(* IEC 61131-3 sources: llm-plc-st-eval/data/definitivo/gpt-4o-2024-08-06/I8/few_shot, 3 files *)

(* ---- ejec_1.st ---- *)
```pascal
FUNCTION_BLOCK FB_Compresor
VAR_INPUT
    pOilOk : BOOL; (* Presión de aceite correcta *)
    tempOk : BOOL; (* Temperatura correcta *)
    sinAlm : BOOL; (* Ausencia de alarmas *)
    btnMarcha : BOOL; (* Botón de marcha *)
    btnParo : BOOL; (* Botón de paro *)
END_VAR
VAR_OUTPUT
    comp : BOOL; (* Compresor en marcha *)
    causaBloqueo : INT; (* Causa de bloqueo *)
END_VAR
VAR
    pOilOkTimer : TON; (* Temporizador para presión de aceite *)
    btnMarchaMem : BOOL; (* Memoria del estado del botón de marcha *)
    btnMarchaRising : BOOL; (* Detección de flanco ascendente del botón de marcha *)
END_VAR

(* Detección de flanco ascendente del botón de marcha *)
btnMarchaRising := btnMarcha AND NOT btnMarchaMem;
btnMarchaMem := btnMarcha;

(* Temporizador para verificar presión de aceite durante 3 segundos continuos *)
pOilOkTimer(IN := pOilOk, PT := T#3S);

(* Determinación de la causa de bloqueo *)
IF NOT pOilOkTimer.Q THEN
    causaBloqueo := 1; (* Falta presión de aceite *)
ELSIF NOT tempOk THEN
    causaBloqueo := 2; (* Falta temperatura correcta *)
ELSIF NOT sinAlm THEN
    causaBloqueo := 3; (* Alarma activa *)
ELSE
    causaBloqueo := 0; (* Ningún bloqueo *)
END_IF

(* Lógica de control del compresor *)
IF btnParo THEN
    comp := FALSE; (* Parar compresor si se pulsa el botón de paro *)
ELSIF comp THEN
    IF causaBloqueo <> 0 THEN
        comp := FALSE; (* Parar compresor si se pierde algún permisivo *)
    END_IF
ELSE
    IF btnMarchaRising AND (causaBloqueo = 0) THEN
        comp := TRUE; (* Arrancar compresor si se pulsa el botón de marcha y no hay bloqueos *)
    END_IF
END_IF

END_FUNCTION_BLOCK
```

(* ---- ejec_2.st ---- *)
```pascal
FUNCTION_BLOCK FB_Compresor
VAR_INPUT
    pOilOk : BOOL; (* Presion de aceite correcta *)
    tempOk : BOOL; (* Temperatura correcta *)
    sinAlm : BOOL; (* Ausencia de alarmas *)
    btnMarcha : BOOL; (* Boton de marcha *)
    btnParo : BOOL; (* Boton de paro *)
END_VAR
VAR_OUTPUT
    comp : BOOL; (* Compresor en marcha *)
    causaBloqueo : INT; (* Causa de bloqueo *)
END_VAR
VAR
    pOilOkTimer : TON; (* Temporizador para presion de aceite *)
    btnMarchaMem : BOOL; (* Memoria de estado del boton de marcha *)
    permisivosOk : BOOL; (* Todos los permisivos estan activos *)
END_VAR

(* Temporizador para verificar presion de aceite durante 3 segundos *)
pOilOkTimer(IN := pOilOk, PT := T#3S);

(* Verificar si todos los permisivos estan activos *)
permisivosOk := pOilOkTimer.Q AND tempOk AND sinAlm;

(* Logica de arranque y paro del compresor *)
IF btnParo THEN
    comp := FALSE; (* Parar compresor si se pulsa btnParo *)
ELSIF NOT comp AND NOT btnMarchaMem AND btnMarcha AND permisivosOk THEN
    comp := TRUE; (* Arrancar compresor si se pulsa btnMarcha y permisivos estan activos *)
END_IF

(* Actualizar memoria del estado del boton de marcha *)
btnMarchaMem := btnMarcha;

(* Determinar la causa de bloqueo *)
IF NOT pOilOk THEN
    causaBloqueo := 1; (* Bloqueo por presion de aceite *)
ELSIF NOT tempOk THEN
    causaBloqueo := 2; (* Bloqueo por temperatura *)
ELSIF NOT sinAlm THEN
    causaBloqueo := 3; (* Bloqueo por alarma activa *)
ELSE
    causaBloqueo := 0; (* No hay bloqueo *)
END_IF
END_FUNCTION_BLOCK
```

(* ---- ejec_3.st ---- *)
```pascal
FUNCTION_BLOCK FB_Compresor
VAR_INPUT
    pOilOk : BOOL; (* Presion de aceite correcta *)
    tempOk : BOOL; (* Temperatura correcta *)
    sinAlm : BOOL; (* Ausencia de alarmas *)
    btnMarcha : BOOL; (* Boton de marcha *)
    btnParo : BOOL; (* Boton de paro *)
END_VAR
VAR_OUTPUT
    comp : BOOL; (* Compresor en marcha *)
    causaBloqueo : INT; (* Causa del bloqueo *)
END_VAR
VAR
    pOilOkTimer : TON; (* Temporizador para presion de aceite *)
    btnMarchaRising : R_TRIG; (* Detector de flanco ascendente para btnMarcha *)
END_VAR

(* Evaluar el flanco ascendente de btnMarcha *)
btnMarchaRising(CLK := btnMarcha);

(* Temporizador para verificar que pOilOk este activo durante 3 segundos continuos *)
pOilOkTimer(IN := pOilOk, PT := T#3S);

(* Determinar la causa del bloqueo *)
IF NOT pOilOk THEN
    causaBloqueo := 1;
ELSIF NOT tempOk THEN
    causaBloqueo := 2;
ELSIF NOT sinAlm THEN
    causaBloqueo := 3;
ELSE
    causaBloqueo := 0;
END_IF

(* Logica de control del compresor *)
IF btnParo THEN
    comp := FALSE; (* Prioridad al boton de paro *)
ELSIF comp THEN
    (* Mantener el compresor en marcha si todos los permisivos se cumplen *)
    IF NOT (pOilOkTimer.Q AND tempOk AND sinAlm) THEN
        comp := FALSE; (* Detener si algun permisivo se pierde *)
    END_IF
ELSE
    (* Arrancar el compresor si se presiona btnMarcha y todos los permisivos se cumplen *)
    IF btnMarchaRising.Q AND pOilOkTimer.Q AND tempOk AND sinAlm THEN
        comp := TRUE;
    END_IF
END_IF
END_FUNCTION_BLOCK
```
